(* IEC 61131-3 sources: llm-plc-st-eval/data/processed_definitivo/qwen2.5-coder_14b/B4/few_shot, 3 files *)

(* ---- ejec_1.st ---- *)
FUNCTION_BLOCK FB_Giro
VAR_INPUT
    btnFwd : BOOL; (* Boton para girar en sentido horario *)
    btnRev : BOOL; (* Boton para girar en sentido antihorario *)
    btnParo : BOOL; (* Boton para parar *)
END_VAR
VAR_OUTPUT
    fwd : BOOL; (* Sentido horario *)
    rev : BOOL; (* Sentido antihorario *)
END_VAR
VAR
    estado : INT := 0; (* Estado actual del sistema *)
    parado : BOOL := TRUE; (* Indica si el motor está parado *)
END_VAR

(* Estado 0: Parado *)
IF btnParo THEN
    estado := 0;
    parado := TRUE;
    fwd := FALSE;
    rev := FALSE;
ELSIF parado AND btnFwd THEN
    estado := 1;
    parado := FALSE;
    fwd := TRUE;
    rev := FALSE;
ELSIF parado AND btnRev THEN
    estado := 2;
    parado := FALSE;
    fwd := FALSE;
    rev := TRUE;
END_IF

(* Estado 1: Girando en sentido horario *)
IF btnParo THEN
    estado := 0;
    parado := TRUE;
    fwd := FALSE;
    rev := FALSE;
ELSIF btnRev THEN
    estado := 2;
    fwd := FALSE;
    rev := TRUE;
END_IF

(* Estado 2: Girando en sentido antihorario *)
IF btnParo THEN
    estado := 0;
    parado := TRUE;
    fwd := FALSE;
    rev := FALSE;
ELSIF btnFwd THEN
    estado := 1;
    fwd := TRUE;
    rev := FALSE;
END_IF

END_FUNCTION_BLOCK

(* ---- ejec_2.st ---- *)
FUNCTION_BLOCK FB_Giro
VAR_INPUT
    btnFwd : BOOL; (* Boton para giro horario *)
    btnRev : BOOL; (* Boton para giro antihorario *)
    btnParo : BOOL; (* Boton para paro *)
END_VAR
VAR_OUTPUT
    fwd : BOOL; (* Giro horario *)
    rev : BOOL; (* Giro antihorario *)
END_VAR
VAR
    estado : INT := 0; (* Estado actual del sistema *)
END_VAR

(* Máquina de estados para controlar el giro del motor *)
CASE estado OF
    0: (* Estado de paro *)
        IF btnFwd THEN
            estado := 1; (* Transición a giro horario *)
        ELSIF btnRev THEN
            estado := 2; (* Transición a giro antihorario *)
        END_IF;
    1: (* Estado de giro horario *)
        fwd := TRUE;
        rev := FALSE;
        IF btnParo THEN
            estado := 0; (* Transición a paro *)
        ELSIF btnRev THEN
            estado := 2; (* Transición a giro antihorario *)
        END_IF;
    2: (* Estado de giro antihorario *)
        fwd := FALSE;
        rev := TRUE;
        IF btnParo THEN
            estado := 0; (* Transición a paro *)
        ELSIF btnFwd THEN
            estado := 1; (* Transición a giro horario *)
        END_IF;
END_CASE;
END_FUNCTION_BLOCK

(* ---- ejec_3.st ---- *)
FUNCTION_BLOCK FB_Giro
VAR_INPUT
    btnFwd : BOOL; (* Boton para girar en sentido horario *)
    btnRev : BOOL; (* Boton para girar en sentido antihorario *)
    btnParo : BOOL; (* Boton para parar el motor *)
END_VAR
VAR_OUTPUT
    fwd : BOOL; (* Salida para giro horario *)
    rev : BOOL; (* Salida para giro antihorario *)
END_VAR
VAR
    estado : INT := 0; (* Estado actual del motor *)
END_VAR

(* Estados: 0 - Parado, 1 - Giro horario, 2 - Giro antihorario *)
CASE estado OF
    0: (* Parado *)
        IF btnFwd THEN
            estado := 1;
        ELSIF btnRev THEN
            estado := 2;
        END_IF;
    1: (* Giro horario *)
        fwd := TRUE;
        rev := FALSE;
        IF btnParo THEN
            estado := 0;
        ELSIF btnRev THEN
            estado := 2;
        END_IF;
    2: (* Giro antihorario *)
        fwd := FALSE;
        rev := TRUE;
        IF btnParo THEN
            estado := 0;
        ELSIF btnFwd THEN
            estado := 1;
        END_IF;
END_CASE;
END_FUNCTION_BLOCK
